// TIA Portal V21 export
// export: Created 2026-11-07T00:00:00Z, ExportSetting WithDefaults
TagTable "Proto tags"
  P_SwOn : Bool  (PLC tag HMI_IF.SwOn, HMI_Connection_1, 100 ms)
